Fanuc KAREL source: KA00117.KL

PROGRAM KA00117
%NOLOCKGROUP
VAR
  SRC: CONFIG
  DST: VECTOR
BEGIN
  SRC.CFG_FLIP = TRUE
  DST = SRC
END KA00117
